(* IEC 61131-3 sources: sis-interlock-demo/src/POUs/Sis/F_SisNe43Valid, 1 file *)

(* ---- F_SisNe43Valid.decl.st ---- *)
// Назначение: достоверность тока 4–20 мА по NAMUR NE 43: 3,6 мА < I < 21,0 мА и значение конечно
//             (пороги — константы PL.GVL_Const, сверить с NE 43). Ток вне диапазона измерения
//             (3,6–3,8 и 20,5–21,0 мА) достоверен: датчик в насыщении показывает выход за шкалу.
// Автор:      kr0nsch
// Версия:     0.1.0
// Документ:   docs/DESIGN.md, раздел «8.3 Аналоговые входы 4–20 мА (NE 43)»
// ВНИМАНИЕ:   код демонстрационный и не предназначен для систем безопасности. Реальная ПАЗ
//             требует определения SIL, сертифицированных аппаратных и программных средств
//             и валидации по ГОСТ Р МЭК 61511.
FUNCTION F_SisNe43Valid : BOOL
VAR_INPUT
    rIn_mA : REAL;   // ток канала, мА
END_VAR
